(* IEC 61131-3 sources: volt/packages/volt-lsp-iec/test-corpus/lenze-mid/Device/Plc Logic/Application/Library Manager/CAA CANopen Stack, 21 files *)

(* ---- BUSSTATE.dut ---- *)
TYPE BUSSTATE :
(
	UNKNOWN,
	ERR_FREE,
	ACTIVE,
	WARNING,
	PASSIVE,
	BUSOFF
);
END_TYPE

(* ---- CANOPEN_KERNEL_ERROR.dut ---- *)
TYPE CANOPEN_KERNEL_ERROR :
(
	CANOPEN_KERNEL_NO_ERROR := 16#0,
	CANOPEN_KERNEL_OTHER_ERROR := 16#1,
	CANOPEN_KERNEL_DATA_OVERFLOW := 16#2,
	CANOPEN_KERNEL_TIMEOUT := 16#3,
	CANOPEN_KERNEL_CANBUS_OFF := 16#10,
	CANOPEN_KERNEL_CAN_ERROR_PASSIVE := 16#11,
	CANOPEN_INTERNAL_FB_ERROR := 16#21,
	CANOPEN_NO_MORE_MEMORY := 16#22,
	CANOPEN_WRONG_PARAMETER := 16#23,
	CANOPEN_NODEID_UNKNOWN := 16#24,
	CANOPEN_NETID_UNKNOWN := 16#25,
	CANOPEN_REQUEST_ERROR := 16#26,
	CANOPEN_SDOCHANNEL_UNKNOWN := 16#27,
	CANOPEN_NO_DRIVER := 16#28,
	CANOPEN_CONFIGURATION_ERROR := 16#29,
	CANOPEN_GUARDING_ERROR := 16#2A
);
END_TYPE

(* ---- DEVICE_STATE.dut ---- *)
TYPE DEVICE_STATE :
(
	INIT,
	RESET_COMM,
	RESET_APP,
	PRE_OPERATIONAL,
	STOPPED,
	OPERATIONAL,
	UNKNOWN,
	NOT_AVAIL
);
END_TYPE

(* ---- EMCY_DATA.dut ---- *)
TYPE EMCY_DATA :
STRUCT
	DEVICE : USINT;
	ABYDUMMY : ARRAY [0..2] OF BYTE;
END_STRUCT
END_TYPE

(* ---- EMCY_ERROR.dut ---- *)
TYPE EMCY_ERROR :
STRUCT
	EMCY_ERROR_CODE : WORD;
	ERROR_REGISTER : BYTE;
	BYDUMMY : BYTE;
	ERROR_FIELD : ARRAY [1..5] OF BYTE;
END_STRUCT
END_TYPE

(* ---- ERROR.dut ---- *)
TYPE ERROR :
(
	NO_ERROR := 0,
	FIRST_ERROR := 10400,
	TIME_OUT := 10401,
	NOT_OPEN := 10404,
	ALREADY_OPEN := 10405,
	ALREADY_CLOSE := 10406,
	REQUEST_ERROR := 10407,
	WRONG_PARAMETER := 10408,
	NODEID_UNKNOWN := 10409,
	SDOCHANNEL_UNKNOWN := 10410,
	INTERNAL_ERROR := 10411,
	NOT_ENOUGH_MEMORY := 10412,
	ABORT_BY_SERVER := 10413,
	INVALID_SEQUENCE_NUMBER := 10414,
	INVALID_BLOCKSIZE := 10415,
	CRC_ERROR := 10416,
	FIRST_MF := 10450,
	LAST_ERROR := 10499
);
END_TYPE

(* ---- NET_INFO.dut ---- *)
TYPE NET_INFO :
STRUCT
	USINETID : USINT;
	UIBAUDRATE : UINT;
	ESTATE : BUSSTATE;
END_STRUCT
END_TYPE

(* ---- PROC_CMD.dut ---- *)
TYPE PROC_CMD :
(
	NONE,
	EXECUTE,
	ABORT
);
END_TYPE

(* ---- PROC_STATE.dut ---- *)
TYPE PROC_STATE :
(
	DORMANT,
	BUSY,
	DONE,
	ABORTED,
	ERROR
);
END_TYPE

(* ---- SDO_ABORT.dut ---- *)
TYPE SDO_ABORT :
STRUCT
END_STRUCT
END_TYPE

(* ---- SDO_MODE.dut ---- *)
TYPE SDO_MODE :
(
	AUTO,
	EXPEDITED,
	SEGMENTED,
	BLOCK
);
END_TYPE

(* ---- SDO_READ.dut ---- *)
TYPE SDO_READ :
STRUCT
	USINODEID : USINT;
	USICHANNEL : USINT;
	UIINDEX : UINT;
	USISUBINDEX : USINT;
	XUSESPECIFICTIMEOUT : BOOL;
	XBLOCKTRANSFER : BOOL;
	USIPST : USINT;
	UISTATE : UINT;
	XLEGACYCRC : BOOL;
	XDUMMY : BOOL;
	UDISIZE : UDINT;
	PDATA : CAA.PVOID;
	UDIABORTCODE : UDINT;
	HDRIVER : CAA.HANDLE;
	HRECEIVER : CAA.HANDLE;
	UDIRXID : UDINT;
	UDITXID : UDINT;
	UDISEGLEN : UDINT;
	UDICURPOS : UDINT;
	TKCURRENTTICK : CAA.TICK;
	XTIMEOUT : BOOL;
	USISEQCNT : USINT;
	UISDOSTATE : UINT;
	TKTIMEOUT : CAA.TICK;
	CTTIMEOUT : CAA.COUNT;
END_STRUCT
END_TYPE

(* ---- SDO_WRITE.dut ---- *)
TYPE SDO_WRITE :
STRUCT
	USINODEID : USINT;
	USICHANNEL : USINT;
	UIINDEX : UINT;
	USISUBINDEX : USINT;
	XUSESPECIFICTIMEOUT : BOOL;
	EMODE : SDO_MODE;
	UISTATE : UINT;
	XLEGACYCRC : BOOL;
	XDUMMY : BOOL;
	UDISIZE : UDINT;
	PDATA : CAA.PVOID;
	UDIABORTCODE : UDINT;
	HDRIVER : CAA.HANDLE;
	HRECEIVER : CAA.HANDLE;
	UDIRXID : UDINT;
	UDITXID : UDINT;
	UDISEQCNT : UDINT;
	UDICURPOS : UDINT;
	TKCURRENTTICK : CAA.TICK;
	XTIMEOUT : BOOL;
	USIBLKSIZE : USINT;
	UISDOSTATE : UINT;
	TKTIMEOUT : CAA.TICK;
	CTTIMEOUT : CAA.COUNT;
END_STRUCT
END_TYPE

(* ---- STK_INFO.dut ---- *)
TYPE STK_INFO :
STRUCT
	USINODEID : USINT;
	ESTATE : STK_STATE;
	ESPEC : STK_SPEC;
END_STRUCT
END_TYPE

(* ---- STK_NODES.dut ---- *)
TYPE STK_NODES :
(
	UNKNOWN := 16#FF,
	LOCAL := 16#0,
	NMT_MASTER := 16#F0,
	CFG_MANAGER := 16#F1,
	SYNC_PRODUCER := 16#F2,
	TIME_PRODUCER := 16#F3
);
END_TYPE

(* ---- STK_SPEC.dut ---- *)
TYPE STK_SPEC :
(
	UNDEFINED := 16#0,
	NMT_SLAVE := 16#1,
	NMT_MASTER := 16#2,
	NMT_FLYMST := 16#4,
	SDO_MANAGER := 16#8,
	CFG_MANAGER := 16#10,
	SYNC_CONSUMER := 16#20,
	SYNC_PRODUCER := 16#40,
	TIME_PRODUCER := 16#80,
	TIME_CONSUMER := 16#100
);
END_TYPE

(* ---- STK_STATE.dut ---- *)
TYPE STK_STATE :
(
	NO_STATE,
	INITALISATION,
	RESET_APPLICATION,
	RESET_COMMUNICATION,
	PRE_OPERATIONAL,
	OPERATIONAL,
	STOPPED
);
END_TYPE

(* ---- OBJECTDICTIONARY.gvl ---- *)
VAR_GLOBAL
	GC_UISTATE_IDX : UINT := 16#1F82;
	GC_UICANOPEN_KERNEL_STATE_IDX : UINT := 16#2001;
	GC_USICANOPEN_KERNEL_STATE_SUBIDX : USINT := 1;
	GC_UIEMCY_DEV_IDX : UINT := 16#2002;
	GC_UIEMCY_IDX : UINT := 16#2003;
	GC_UIEMCY_SUBIDX : USINT := 1;
	GC_UIPERMITSDOTRANSMISSION_IDX : UINT := 16#2004;
	GC_UISDOCHANNELLIMIT_IDX : UINT := 16#2005;
	GC_UIBLOCKFDTACCESS_IDX : UINT := 16#2006;
END_VAR

(* ---- VERSIONCONSTANTS.gvl ---- *)
VAR_GLOBAL
	GC_BYVERSION : BYTE := 1;
	GC_BYVERSION_1 : BYTE := 0;
END_VAR

(* ---- ICANOPENSTACK.itf ---- *)
INTERFACE ICANOPENSTACK
END_INTERFACE

METHOD SDOABORT : PROC_STATE
VAR_INPUT
	ECMD : PROC_CMD;
	PPARAM : POINTER TO SDO_ABORT;
END_VAR
VAR_OUTPUT
	EERROR : ERROR;
END_VAR
END_METHOD

METHOD SDOWRITE : PROC_STATE
VAR_INPUT
	ECMD : PROC_CMD;
	PPARAM : POINTER TO SDO_WRITE;
END_VAR
VAR_OUTPUT
	EERROR : ERROR;
END_VAR
END_METHOD

METHOD SDOREAD : PROC_STATE
VAR_INPUT
	ECMD : PROC_CMD;
	PPARAM : POINTER TO SDO_READ;
END_VAR
VAR_OUTPUT
	EERROR : ERROR;
END_VAR
END_METHOD

METHOD STKOPEN : PROC_STATE
VAR_INPUT
	ECMD : PROC_CMD;
	USINETID : USINT;
	USINODEID : USINT;
	UIBAUDRATE : UINT;
	ESPEC : STK_SPEC;
END_VAR
VAR_OUTPUT
	EERROR : ERROR;
END_VAR
END_METHOD

METHOD STKCLOSE : PROC_STATE
VAR_INPUT
	ECMD : PROC_CMD;
END_VAR
VAR_OUTPUT
	EERROR : ERROR;
END_VAR
END_METHOD

METHOD STKGETINFO : PROC_STATE
VAR_INPUT
	ECMD : PROC_CMD;
	PSTKINFO : POINTER TO STK_INFO;
	PNETINFO : POINTER TO NET_INFO;
END_VAR
VAR_OUTPUT
	EERROR : ERROR;
END_VAR
END_METHOD

(* ---- GETSUPPLIERVERSION.pou ---- *)
FUNCTION GETSUPPLIERVERSION : WORD
VAR_INPUT
	XDUMMY : BOOL;
END_VAR
END_FUNCTION
